Fanuc KAREL source: ko00106.KL

-- PROVISIONAL review KL for V770-1; original PC SHA256 81e7323237f620edaf3aed086c5b9a278b2b022823a6dd13e95aec8148650965
-- Incomplete behavior may be omitted. Consult companion uncertainty JSON. Do not deploy.
PROGRAM KO00106
%NOLOCKGROUP
VAR
  A : REAL
  B : INTEGER
  OUT : REAL
BEGIN
  -- UNRESOLVED_PC offsets 5-13; opcodes 9D,64,23
  -- UNRESOLVED_PC offsets 18-29; opcodes 2E,23
  -- UNRESOLVED_PC offsets 34-57; opcodes 27,22,27,21,64,76,23
  -- UNRESOLVED_PC offsets 62-66; opcodes 7F
END KO00106
